Fanuc KAREL source: KT00512.KL

PROGRAM KT00512
%NOLOCKGROUP
VAR
  P1: XYZWPR
  P2: JOINTPOS
  OUT: JOINTPOS
BEGIN
  P1.X = 1.0
  OUT = P1 : P2
END KT00512
